// TIA Portal V20 export
// export: Created 2026-10-19T18:45:34.7281503Z, ExportSetting None, DisplayName Totally Integrated Automation Portal, DisplayVersion V20 Update 6, DisplayName TIA Portal Openness, DisplayVersion V20 Update 6, DisplayName TIA Portal Version Control Interface, DisplayVersion V20 Update 6, DisplayName SINAMICS Startdrive Advanced, DisplayVersion V20 SP1, DisplayName SINAMICS Startdrive G130, G150, S120, S150, SINAMICS MV, G220, S200, S210, DisplayVersion V20 SP1, DisplayName SINAMICS Startdrive G110M, G120, G120C, G120D, G120P, G115D, DisplayVersion V20 SP1, DisplayName STEP 7 Professional, DisplayVersion V20 Update 6, DisplayName STEP 7 Safety, DisplayVersion V20 Update 2, DisplayName WinCC Basic/Comfort/Advanced, DisplayVersion V20 Update 6, DisplayName WinCC Unified, DisplayVersion V20 Update 6
VAR_GLOBAL   // PLC tag table "IO_VFDs_2"
   C2104_ActualTorque AT %IW570 : Word;
   C2102_ActualSpeed AT %IW538 : Word;
   C2202_Inputs AT %IW622 : Word;
   C2205_ActualTorque AT %IW762 : Word;
   C2206_ActualTorque AT %IW778 : Word;
   C2202_StatusWord AT %IW612 : Word;
   C2103_ActualTorque AT %IW554 : Word;
   C2105_ActualTorque AT %IW586 : Word;
   C2105_ControlWord AT %QW236 : Word;
   VTD2_ActualTorque AT %IW505 : Word;
   C2202_ActualSpeed AT %IW614 : Word;
   C2202_ActualTorque AT %IW618 : Word;
   C2103_ActualSpeed AT %IW550 : Word;
   VTD2_AccFactor AT %QW1517 : Word;
   C2206_Inputs AT %IW782 : Word;
   C2106_Inputs AT %IW606 : Word;
   C2104_Inputs AT %IW574 : Word;
   C2106_StatusWord AT %IW596 : Word;
   C2205_Inputs AT %IW766 : Word;
   C2204_ActualCurrent AT %IW744 : Word;
   C2202_ActualCurrent AT %IW616 : Word;
   C2203_ActualSpeed AT %IW630 : Word;
   C2205_ActualSpeed AT %IW758 : Word;
   C2105_StatusWord AT %IW580 : Word;
   C2105_ActualCurrent AT %IW584 : Word;
   C2102_ActualCurrent AT %IW540 : Word;
   C2104_StatusWord AT %IW564 : Word;
   C2204_ControlWord AT %QW268 : Word;
   C2204_Inputs AT %IW750 : Word;
   VTD2_ControlWord AT %QW216 : Word;
   C2206_ControlWord AT %QW284 : Word;
   CVTD2_ActualCurrent AT %IW515 : Word;
   C2103_StatusWord AT %IW548 : Word;
   C2206_ActualCurrent AT %IW776 : Word;
   C2103_Inputs AT %IW558 : Word;
   C2204_ActualTorque AT %IW746 : Word;
   C2204_ActualSpeed AT %IW742 : Word;
   C2105_ActualSpeed AT %IW582 : Word;
   C2203_StatusWord AT %IW628 : Word;
   VTD2_StatusWord AT %IW499 : Word;
   C2106_ActualSpeed AT %IW598 : Word;
   CVTD2_ControlWord AT %QW184 : Word;
   CVTD2_StatusWord AT %IW511 : Word;
   C2106_ActualTorque AT %IW602 : Word;
   C2104_ActualCurrent AT %IW568 : Word;
   C2103_ControlWord AT %QW220 : Word;
   C2102_ControlWord AT %QW198 : Word;
   C2205_ControlWord AT %QW276 : Word;
   CVTD2_Inputs AT %IW521 : Word;
   C2105_Inputs AT %IW590 : Word;
   C2104_ControlWord AT %QW228 : Word;
   C2203_ActualCurrent AT %IW632 : Word;
   VTD2_ActualSpeed AT %IW501 : Word;
   C2203_ControlWord AT %QW260 : Word;
   C2205_ActualCurrent AT %IW760 : Word;
   CVTD2_ActualTorque AT %IW517 : Word;
   C2102_StatusWord AT %IW536 : Word;
   C2102_ActualTorque AT %IW542 : Word;
   C2106_ActualCurrent AT %IW600 : Word;
   CVTD2_ActualSpeed AT %IW513 : Word;
   C2203_ActualTorque AT %IW634 : Word;
   CVTD2_MainSetpoint AT %QW186 : Word;
   C2102_Inputs AT %IW546 : Word;
   C2104_ActualSpeed AT %IW566 : Word;
   C2203_Inputs AT %IW638 : Word;
   C2205_StatusWord AT %IW756 : Word;
   C2202_ControlWord AT %QW252 : Word;
   C2206_StatusWord AT %IW772 : Word;
   C2103_ActualCurrent AT %IW552 : Word;
   VTD2_ActualCurrent AT %IW503 : Word;
   C2106_ControlWord AT %QW244 : Word;
   C2206_ActualSpeed AT %IW774 : Word;
   C2204_StatusWord AT %IW740 : Word;
END_VAR
